(* IEC 61131-3 sources: codesys-framework/txt/application/ToDo/Hardware/IO/Cylinder/FB_Cylinder, 1 file *)

(* ---- Reset.method.st ---- *)
METHOD Reset : BOOL
VAR_INPUT
END_VAR

// --- BEGIN IMPLEMENTATION ---

SUPER^.Reset();

Reset := TRUE;
